// TIA Portal V20 export
// export: Created 2026-10-19T18:06:18.2529775Z, ExportSetting WithDefaults, DisplayName Totally Integrated Automation Portal, DisplayVersion V20 Update 6, DisplayName TIA Portal Openness, DisplayVersion V20 Update 6, DisplayName TIA Portal Version Control Interface, DisplayVersion V20 Update 6, DisplayName SINAMICS Startdrive Advanced, DisplayVersion V20 SP1, DisplayName SINAMICS Startdrive G130, G150, S120, S150, SINAMICS MV, G220, S200, S210, DisplayVersion V20 SP1, DisplayName SINAMICS Startdrive G110M, G120, G120C, G120D, G120P, G115D, DisplayVersion V20 SP1, DisplayName STEP 7 Professional, DisplayVersion V20 Update 6, DisplayName STEP 7 Safety, DisplayVersion V20 Update 2, DisplayName WinCC Basic/Comfort/Advanced, DisplayVersion V20 Update 6, DisplayName WinCC Unified, DisplayVersion V20 Update 6
FUNCTION_BLOCK "SAI_Cyclic_WeightProc"   // FB29, LAD
TITLE = Cyclic Weighing Process: Send PLC commands and read Weight data and device status bits
{ S7_Optimized_Access := 'FALSE' }
VERSION : 0.1
// stored: AutoNumber true, IsIECCheckEnabled false, SetENOAutomatically false, UDAEnableTagReadback false
   VAR_INPUT
      WeightCmd { ExternalAccessible := 'False'; ExternalVisible := 'False'; ExternalWritable := 'False'} : Word := 3;
      MB_DevStatus : Word;
   END_VAR
   VAR_OUTPUT
      RealTimeWeight { ExternalVisible := 'False'; ExternalWritable := 'False'} : Real;
      StableWeight { ExternalVisible := 'False'; ExternalWritable := 'False'} : Real;
      DataOK : Bool;
      Motion : Bool;
      NetMode : Bool;
      Alarm : Bool;
      Done { ExternalAccessible := 'False'; ExternalVisible := 'False'; ExternalWritable := 'False'} : Bool;
      Error { ExternalAccessible := 'False'; ExternalVisible := 'False'; ExternalWritable := 'False'} : Bool;
   END_VAR
   VAR_IN_OUT
      TareImmediate { ExternalAccessible := 'False'; ExternalVisible := 'False'; ExternalWritable := 'False'} : Bool;
      TareStable { ExternalAccessible := 'False'; ExternalVisible := 'False'; ExternalWritable := 'False'} : Bool;
      ZeroImmediate { ExternalAccessible := 'False'; ExternalVisible := 'False'; ExternalWritable := 'False'} : Bool;
      ZeroStable { ExternalAccessible := 'False'; ExternalVisible := 'False'; ExternalWritable := 'False'} : Bool;
      PreTareValue : Real;
      PreTare : Bool;
      ClearTare { ExternalAccessible := 'False'; ExternalVisible := 'False'; ExternalWritable := 'False'} : Bool;
      MB_Value : Real;
      MB_Response : Word;
      MB_CmdValue : Real;
      MB_Command : Word;
   END_VAR
   VAR DB_SPECIFIC
      WriteTrigger { ExternalAccessible := 'False'; ExternalVisible := 'False'; ExternalWritable := 'False'} : Bool;
      RestoreTrigger { ExternalAccessible := 'False'; ExternalVisible := 'False'; ExternalWritable := 'False'} : Bool;
      Cmd { ExternalAccessible := 'False'; ExternalVisible := 'False'; ExternalWritable := 'False'} : Int;
      TareStablePTrigger : Bool;
      ZeroStablePTrigger : Bool;
      ZeroImmedTrigger : Bool;
      TareImmedTrigger : Bool;
      ClearTareTrigger : Bool;
      PreTareTrigger : Bool;
   END_VAR
   VAR_TEMP
      DevStatus : "SAI_MB_DeviceStatus";
   END_VAR
   VAR_TEMP   // added for the SCL form of the ladder/FBD networks
      _w1 : Bool;
   END_VAR
BEGIN

REGION Network 1: During 1st PLC scan, moves the default weight reporting command to the cyclic command output word
   // During 1st scan, moves the default weight reporting command to the cyclic command output word
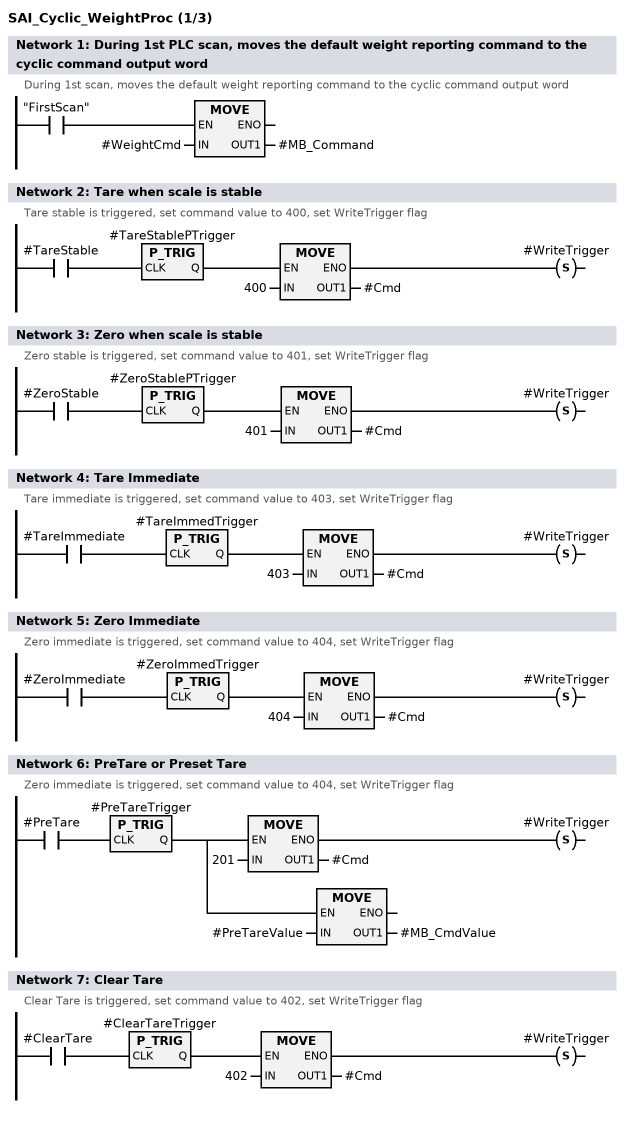
   RUNG wire#powerrail
      Contact( "FirstScan" )
      { S7_GenerateENO := "TRUE" } Move(in := #WeightCmd, out1 => #MB_Command)
   END_RUNG
   // the same network as SCL:
   IF "FirstScan" THEN #MB_Command := #WeightCmd; END_IF;
END_REGION

REGION Network 2: Tare when scale is stable
   // Tare stable is triggered, set command value to 400, set WriteTrigger flag
   RUNG wire#powerrail
      Contact( #TareStable )
      P_Trig( #TareStablePTrigger )
      { S7_GenerateENO := "TRUE" } Move(in := 400, out1 => #Cmd)
      S_Coil( #WriteTrigger )
   END_RUNG
   // the same network as SCL:
   // ENO of a box is taken as its EN; it also drops when the box reports an error
   #_w1 := #TareStable AND NOT #TareStablePTrigger;   // rising edge
   #TareStablePTrigger := #TareStable;
   IF #_w1 THEN
       #Cmd := 400;
       #WriteTrigger := TRUE;
   END_IF;
END_REGION

REGION Network 3: Zero when scale is stable
   // Zero stable is triggered, set command value to 401, set WriteTrigger flag
   RUNG wire#powerrail
      Contact( #ZeroStable )
      P_Trig( #ZeroStablePTrigger )
      { S7_GenerateENO := "TRUE" } Move(in := 401, out1 => #Cmd)
      S_Coil( #WriteTrigger )
   END_RUNG
   // the same network as SCL:
   // ENO of a box is taken as its EN; it also drops when the box reports an error
   #_w1 := #ZeroStable AND NOT #ZeroStablePTrigger;   // rising edge
   #ZeroStablePTrigger := #ZeroStable;
   IF #_w1 THEN
       #Cmd := 401;
       #WriteTrigger := TRUE;
   END_IF;
END_REGION

REGION Network 4: Tare Immediate
   // Tare immediate is triggered, set command value to 403, set WriteTrigger flag
   RUNG wire#powerrail
      Contact( #TareImmediate )
      P_Trig( #TareImmedTrigger )
      { S7_GenerateENO := "TRUE" } Move(in := 403, out1 => #Cmd)
      S_Coil( #WriteTrigger )
   END_RUNG
   // the same network as SCL:
   // ENO of a box is taken as its EN; it also drops when the box reports an error
   #_w1 := #TareImmediate AND NOT #TareImmedTrigger;   // rising edge
   #TareImmedTrigger := #TareImmediate;
   IF #_w1 THEN
       #Cmd := 403;
       #WriteTrigger := TRUE;
   END_IF;
END_REGION

REGION Network 5: Zero Immediate
   // Zero immediate is triggered, set command value to 404, set WriteTrigger flag
   RUNG wire#powerrail
      Contact( #ZeroImmediate )
      P_Trig( #ZeroImmedTrigger )
      { S7_GenerateENO := "TRUE" } Move(in := 404, out1 => #Cmd)
      S_Coil( #WriteTrigger )
   END_RUNG
   // the same network as SCL:
   // ENO of a box is taken as its EN; it also drops when the box reports an error
   #_w1 := #ZeroImmediate AND NOT #ZeroImmedTrigger;   // rising edge
   #ZeroImmedTrigger := #ZeroImmediate;
   IF #_w1 THEN
       #Cmd := 404;
       #WriteTrigger := TRUE;
   END_IF;
END_REGION

REGION Network 6: PreTare or Preset Tare
   // Zero immediate is triggered, set command value to 404, set WriteTrigger flag
   RUNG wire#powerrail
      Contact( #PreTare )
      P_Trig( #PreTareTrigger )
      wire#w1
      { S7_GenerateENO := "TRUE" } Move(in := 201, out1 => #Cmd)
      S_Coil( #WriteTrigger )
   END_RUNG
   RUNG wire#w1
      { S7_GenerateENO := "TRUE" } Move(in := #PreTareValue, out1 => #MB_CmdValue)
   END_RUNG
   // the same network as SCL:
   // ENO of a box is taken as its EN; it also drops when the box reports an error
   #_w1 := #PreTare AND NOT #PreTareTrigger;   // rising edge
   #PreTareTrigger := #PreTare;
   IF #_w1 THEN
       #Cmd := 201;
       #WriteTrigger := TRUE;
       #MB_CmdValue := #PreTareValue;
   END_IF;
END_REGION

REGION Network 7: Clear Tare
   // Clear Tare is triggered, set command value to 402, set WriteTrigger flag
   RUNG wire#powerrail
      Contact( #ClearTare )
      P_Trig( #ClearTareTrigger )
      { S7_GenerateENO := "TRUE" } Move(in := 402, out1 => #Cmd)
      S_Coil( #WriteTrigger )
   END_RUNG
   // the same network as SCL:
   // ENO of a box is taken as its EN; it also drops when the box reports an error
   #_w1 := #ClearTare AND NOT #ClearTareTrigger;   // rising edge
   #ClearTareTrigger := #ClearTare;
   IF #_w1 THEN
       #Cmd := 402;
       #WriteTrigger := TRUE;
   END_IF;
END_REGION

REGION Network 8: Deliver the command
   // Move the command value to output, reset flags
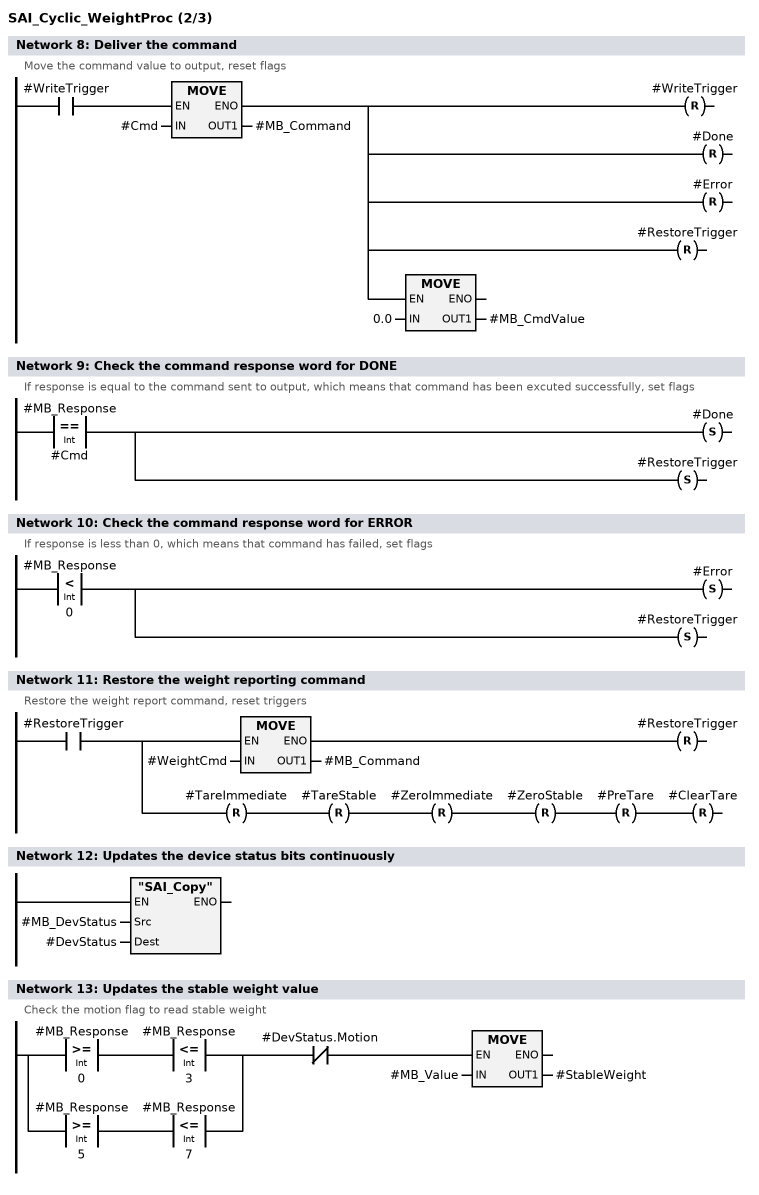
   RUNG wire#powerrail
      Contact( #WriteTrigger )
      { S7_GenerateENO := "TRUE" } Move(in := #Cmd, out1 => #MB_Command)
      wire#w1
      R_Coil( #WriteTrigger )
   END_RUNG
   RUNG wire#w1
      R_Coil( #Done )
   END_RUNG
   RUNG wire#w1
      R_Coil( #Error )
   END_RUNG
   RUNG wire#w1
      R_Coil( #RestoreTrigger )
   END_RUNG
   RUNG wire#w1
      { S7_GenerateENO := "TRUE" } Move(in := 0.0, out1 => #MB_CmdValue)
   END_RUNG
   // the same network as SCL:
   // ENO of a box is taken as its EN; it also drops when the box reports an error
   IF #WriteTrigger THEN #MB_Command := #Cmd; END_IF;
   #_w1 := #WriteTrigger;
   IF #_w1 THEN
       #WriteTrigger := FALSE;
       #Done := FALSE;
       #Error := FALSE;
       #RestoreTrigger := FALSE;
       #MB_CmdValue := 0.0;
   END_IF;
END_REGION

REGION Network 9: Check the command response word for DONE
   // If response is equal to the command sent to output, which means that command has been excuted successfully, set flags
   RUNG wire#powerrail
      { S7_Templates := "SrcType := Int" } EQ_Contact(in1 := #MB_Response, in2 := #Cmd)
      wire#w1
      S_Coil( #Done )
   END_RUNG
   RUNG wire#w1
      S_Coil( #RestoreTrigger )
   END_RUNG
   // the same network as SCL:
   IF #MB_Response = #Cmd THEN
       #Done := TRUE;
       #RestoreTrigger := TRUE;
   END_IF;
END_REGION

REGION Network 10: Check the command response word for ERROR
   // If response is less than 0, which means that command has failed, set flags
   RUNG wire#powerrail
      { S7_Templates := "SrcType := Int" } LT_Contact(in1 := #MB_Response, in2 := 0)
      wire#w1
      S_Coil( #Error )
   END_RUNG
   RUNG wire#w1
      S_Coil( #RestoreTrigger )
   END_RUNG
   // the same network as SCL:
   IF #MB_Response < 0 THEN
       #Error := TRUE;
       #RestoreTrigger := TRUE;
   END_IF;
END_REGION

REGION Network 11: Restore the weight reporting command
   // Restore the weight report command, reset triggers
   RUNG wire#powerrail
      Contact( #RestoreTrigger )
      wire#w1
      { S7_GenerateENO := "TRUE" } Move(in := #WeightCmd, out1 => #MB_Command)
      R_Coil( #RestoreTrigger )
   END_RUNG
   RUNG wire#w1
      R_Coil( #TareImmediate )
      R_Coil( #TareStable )
      R_Coil( #ZeroImmediate )
      R_Coil( #ZeroStable )
      R_Coil( #PreTare )
      R_Coil( #ClearTare )
   END_RUNG
   // the same network as SCL:
   // ENO of a box is taken as its EN; it also drops when the box reports an error
   IF #RestoreTrigger THEN #MB_Command := #WeightCmd; END_IF;
   #_w1 := #RestoreTrigger;
   IF #_w1 THEN
       #RestoreTrigger := FALSE;
       #TareImmediate := FALSE;
       #TareStable := FALSE;
       #ZeroImmediate := FALSE;
       #ZeroStable := FALSE;
       #PreTare := FALSE;
       #ClearTare := FALSE;
   END_IF;
END_REGION

REGION Network 12: Updates the device status bits continuously
   RUNG wire#powerrail
      "SAI_Copy"(Src := #MB_DevStatus, Dest := #DevStatus)
   END_RUNG
   // the same network as SCL:
   "SAI_Copy"(Src := #MB_DevStatus, Dest := #DevStatus);
END_REGION

REGION Network 13: Updates the stable weight value
   // Check the motion flag to read stable weight
   RUNG wire#powerrail
      { S7_Templates := "SrcType := Int" } GE_Contact(in1 := #MB_Response, in2 := 0)
      { S7_Templates := "SrcType := Int" } LE_Contact(in1 := #MB_Response, in2 := 3)
      wire#w1
      I_Contact( #DevStatus.Motion )
      { S7_GenerateENO := "TRUE" } Move(in := #MB_Value, out1 => #StableWeight)
   END_RUNG
   RUNG wire#powerrail
      { S7_Templates := "SrcType := Int" } GE_Contact(in1 := #MB_Response, in2 := 5)
      { S7_Templates := "SrcType := Int" } LE_Contact(in1 := #MB_Response, in2 := 7)
   END_RUNG wire#w1
   // the same network as SCL:
   IF (((#MB_Response >= 0) AND (#MB_Response <= 3)) OR ((#MB_Response >= 5) AND (#MB_Response <= 7))) AND NOT #DevStatus.Motion THEN
       #StableWeight := #MB_Value;
   END_IF;
END_REGION

REGION Network 14: Updates the real time weight value
   // Read real time weight
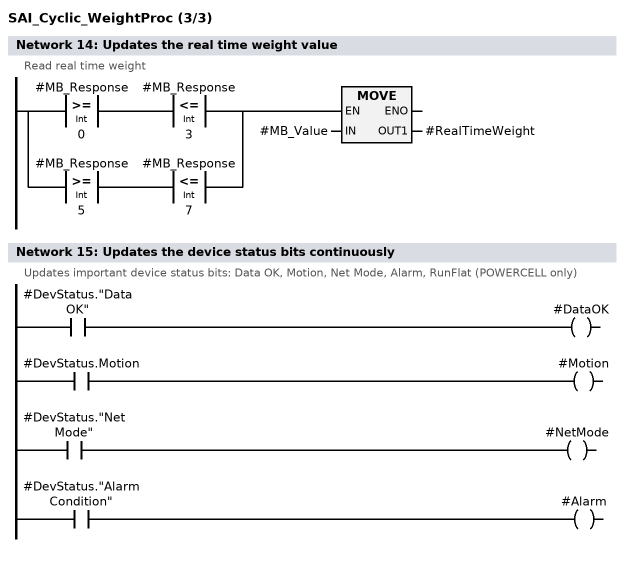
   RUNG wire#powerrail
      { S7_Templates := "SrcType := Int" } GE_Contact(in1 := #MB_Response, in2 := 0)
      { S7_Templates := "SrcType := Int" } LE_Contact(in1 := #MB_Response, in2 := 3)
      wire#w1
      { S7_GenerateENO := "TRUE" } Move(in := #MB_Value, out1 => #RealTimeWeight)
   END_RUNG
   RUNG wire#powerrail
      { S7_Templates := "SrcType := Int" } GE_Contact(in1 := #MB_Response, in2 := 5)
      { S7_Templates := "SrcType := Int" } LE_Contact(in1 := #MB_Response, in2 := 7)
   END_RUNG wire#w1
   // the same network as SCL:
   IF ((#MB_Response >= 0) AND (#MB_Response <= 3)) OR ((#MB_Response >= 5) AND (#MB_Response <= 7)) THEN
       #RealTimeWeight := #MB_Value;
   END_IF;
END_REGION

REGION Network 15: Updates the device status bits continuously
   // Updates important device status bits: Data OK, Motion, Net Mode, Alarm, RunFlat (POWERCELL only)
   RUNG wire#powerrail
      Contact( #DevStatus."Data OK" )
      Coil( #DataOK )
   END_RUNG
   RUNG wire#powerrail
      Contact( #DevStatus.Motion )
      Coil( #Motion )
   END_RUNG
   RUNG wire#powerrail
      Contact( #DevStatus."Net Mode" )
      Coil( #NetMode )
   END_RUNG
   RUNG wire#powerrail
      Contact( #DevStatus."Alarm Condition" )
      Coil( #Alarm )
   END_RUNG
   // the same network as SCL:
   #DataOK := #DevStatus."Data OK";
   #Motion := #DevStatus.Motion;
   #NetMode := #DevStatus."Net Mode";
   #Alarm := #DevStatus."Alarm Condition";
END_REGION
END_FUNCTION_BLOCK
